(* IEC 61131-3 sources: nautilus/examples/it-rack, 2 files *)

(* ---- hw_types.st ---- *)
(*
  Generated by `naut prometheus import`: the IT-hardware UDT set from
  docs/design/it-drivers.md §2. Do not edit — every importer (snmp, redfish,
  prometheus) writes this same file, so re-running any of them restores it.
  Member order is the wire order the drivers deliver; the compiled TYPE
  must match it slot for slot, which is why it is generated and not typed.
*)

TYPE
  CPU : STRUCT
    Model : STRING;
    Cores : DINT;
    Health : DINT;
    Fault : BOOL;
    TempC : REAL;
    Pct : REAL;
  END_STRUCT;
  DIMM : STRUCT
    Locator : STRING;
    CapacityGB : REAL;
    Manufacturer : STRING;
    PartNumber : STRING;
    Health : DINT;
    Fault : BOOL;
    TempC : REAL;
  END_STRUCT;
  Drive : STRUCT
    Bay : DINT;
    Name : STRING;
    Model : STRING;
    Serial : STRING;
    CapacityGB : REAL;
    Protocol : STRING;
    MediaType : STRING;
    Health : DINT;
    Fault : BOOL;
    PredictedFailure : BOOL;
    TempC : REAL;
    Present : BOOL;
  END_STRUCT;
  Fan : STRUCT
    Name : STRING;
    Present : BOOL;
    RPM : REAL;
    Pct : REAL;
    Fault : BOOL;
  END_STRUCT;
  NetPort : STRUCT
    Name : STRING;
    LinkUp : BOOL;
    SpeedGbps : REAL;
    MAC : STRING;
  END_STRUCT;
  PCIeDevice : STRUCT
    Slot : DINT;
    Name : STRING;
    Model : STRING;
    Manufacturer : STRING;
    Firmware : STRING;
    Health : DINT;
    Fault : BOOL;
    Ports : DINT;
    TempC : REAL;
  END_STRUCT;
  PDU : STRUCT
    Online : BOOL;
    Name : STRING;
    Model : STRING;
    Serial : STRING;
    Amps : REAL;
    Watts : REAL;
    Overload : BOOL;
    OutletCount : DINT;
  END_STRUCT;
  PDUOutlet : STRUCT
    Index : DINT;
    Name : STRING;
    On : BOOL;
    Amps : REAL;
    Watts : REAL;
  END_STRUCT;
  PSU : STRUCT
    Name : STRING;
    Present : BOOL;
    Fault : BOOL;
    InputOk : BOOL;
    InputV : REAL;
    OutputW : REAL;
    CapacityW : REAL;
  END_STRUCT;
  Server : STRUCT
    Online : BOOL;
    PowerOn : BOOL;
    Health : DINT;
    Fault : BOOL;
    Warning : BOOL;
    Model : STRING;
    Serial : STRING;
    UptimeS : DINT;
    CpuPct : REAL;
    MemPct : REAL;
    Load1 : REAL;
    RootDiskPct : REAL;
    InletTempC : REAL;
    MaxTempC : REAL;
    PowerW : REAL;
    FanCount : DINT;
    PsuCount : DINT;
    TempCount : DINT;
  END_STRUCT;
  Switch : STRUCT
    Online : BOOL;
    Name : STRING;
    Model : STRING;
    Serial : STRING;
    UptimeS : DINT;
    CpuPct : REAL;
    MemPct : REAL;
    TempC : REAL;
    Fault : BOOL;
    PortsTotal : DINT;
    PortsUp : DINT;
  END_STRUCT;
  SwitchPort : STRUCT
    Index : DINT;
    Name : STRING;
    Alias : STRING;
    AdminUp : BOOL;
    OperUp : BOOL;
    Down : BOOL;
    SpeedMbps : REAL;
    InBps : REAL;
    OutBps : REAL;
    InPct : REAL;
    OutPct : REAL;
    InErrors : DINT;
    OutErrors : DINT;
    InDiscards : DINT;
    OutDiscards : DINT;
    ErrorRate : REAL;
    PoeOn : BOOL;
    PoeW : REAL;
    InBroadcastPps : REAL;
    InMulticastPps : REAL;
  END_STRUCT;
  TempSensor : STRUCT
    Name : STRING;
    Value : REAL;
    Fault : BOOL;
    High : BOOL;
    HighHigh : BOOL;
    HighSP : REAL;
    HighHighSP : REAL;
  END_STRUCT;
  UPS : STRUCT
    Online : BOOL;
    Name : STRING;
    Model : STRING;
    Serial : STRING;
    OnBattery : BOOL;
    LowBattery : BOOL;
    BatteryFault : BOOL;
    Fault : BOOL;
    ChargePct : REAL;
    RuntimeMin : REAL;
    LoadPct : REAL;
    InputV : REAL;
    OutputV : REAL;
    BatteryTempC : REAL;
  END_STRUCT;
END_TYPE

(* ---- rack.st ---- *)
(* rack.st — the rollups a rack needs that no single device carries: how
   many switch ports are up, whether anything in the rack is faulted, and
   the hottest thing in it. Everything else — every port's status, every
   fan's RPM, every sensor's thresholds — is already a UDT tag the drivers
   deliver, alarmed by the rules in nautilus.yaml, so this program stays
   small on purpose.

   Every driver-fed tag is read under its source's __Online companion: a
   device that stops answering keeps its last values (Stale) rather than
   dropping to zero, so the guard is what keeps a dark switch from being
   counted as 24 healthy ports. *)
PROGRAM Rack
VAR_EXTERNAL
  SW1 : Switch;
  SW1_Port01 : SwitchPort; SW1_Port02 : SwitchPort; SW1_Port03 : SwitchPort; SW1_Port04 : SwitchPort;
  SW1_Port05 : SwitchPort; SW1_Port06 : SwitchPort; SW1_Port07 : SwitchPort; SW1_Port08 : SwitchPort;
  SW1_Port09 : SwitchPort; SW1_Port10 : SwitchPort; SW1_Port11 : SwitchPort; SW1_Port12 : SwitchPort;
  SW1_Port13 : SwitchPort; SW1_Port14 : SwitchPort; SW1_Port15 : SwitchPort; SW1_Port16 : SwitchPort;
  SW1_Port17 : SwitchPort; SW1_Port18 : SwitchPort; SW1_Port19 : SwitchPort; SW1_Port20 : SwitchPort;
  SW1_Port21 : SwitchPort; SW1_Port22 : SwitchPort; SW1_Port23 : SwitchPort; SW1_Port24 : SwitchPort;
  SW1_Port25 : SwitchPort; SW1_Port26 : SwitchPort; SW1_Port27 : SwitchPort; SW1_Port28 : SwitchPort;
  SW1__Online : BOOL;
  MIRA1 : Server;
  MIRA1__Online : BOOL;

  PortsUp : INT;
  PortsDown : INT;
  DevicesOnline : INT;
  RackFault : BOOL;
  RackMaxTempC : REAL;
END_VAR
VAR
  up : INT;
  down : INT;
END_VAR

DevicesOnline := 0;
IF SW1__Online THEN DevicesOnline := DevicesOnline + 1; END_IF;
IF MIRA1__Online THEN DevicesOnline := DevicesOnline + 1; END_IF;

(* Ports: up = link; down = enabled but no link (Down is the driver's own
   derived member, AdminUp AND NOT OperUp — a port nobody enabled is
   neither). *)
up := 0; down := 0;
IF SW1__Online THEN
  IF SW1_Port01.OperUp THEN up := up + 1; END_IF; IF SW1_Port01.Down THEN down := down + 1; END_IF;
  IF SW1_Port02.OperUp THEN up := up + 1; END_IF; IF SW1_Port02.Down THEN down := down + 1; END_IF;
  IF SW1_Port03.OperUp THEN up := up + 1; END_IF; IF SW1_Port03.Down THEN down := down + 1; END_IF;
  IF SW1_Port04.OperUp THEN up := up + 1; END_IF; IF SW1_Port04.Down THEN down := down + 1; END_IF;
  IF SW1_Port05.OperUp THEN up := up + 1; END_IF; IF SW1_Port05.Down THEN down := down + 1; END_IF;
  IF SW1_Port06.OperUp THEN up := up + 1; END_IF; IF SW1_Port06.Down THEN down := down + 1; END_IF;
  IF SW1_Port07.OperUp THEN up := up + 1; END_IF; IF SW1_Port07.Down THEN down := down + 1; END_IF;
  IF SW1_Port08.OperUp THEN up := up + 1; END_IF; IF SW1_Port08.Down THEN down := down + 1; END_IF;
  IF SW1_Port09.OperUp THEN up := up + 1; END_IF; IF SW1_Port09.Down THEN down := down + 1; END_IF;
  IF SW1_Port10.OperUp THEN up := up + 1; END_IF; IF SW1_Port10.Down THEN down := down + 1; END_IF;
  IF SW1_Port11.OperUp THEN up := up + 1; END_IF; IF SW1_Port11.Down THEN down := down + 1; END_IF;
  IF SW1_Port12.OperUp THEN up := up + 1; END_IF; IF SW1_Port12.Down THEN down := down + 1; END_IF;
  IF SW1_Port13.OperUp THEN up := up + 1; END_IF; IF SW1_Port13.Down THEN down := down + 1; END_IF;
  IF SW1_Port14.OperUp THEN up := up + 1; END_IF; IF SW1_Port14.Down THEN down := down + 1; END_IF;
  IF SW1_Port15.OperUp THEN up := up + 1; END_IF; IF SW1_Port15.Down THEN down := down + 1; END_IF;
  IF SW1_Port16.OperUp THEN up := up + 1; END_IF; IF SW1_Port16.Down THEN down := down + 1; END_IF;
  IF SW1_Port17.OperUp THEN up := up + 1; END_IF; IF SW1_Port17.Down THEN down := down + 1; END_IF;
  IF SW1_Port18.OperUp THEN up := up + 1; END_IF; IF SW1_Port18.Down THEN down := down + 1; END_IF;
  IF SW1_Port19.OperUp THEN up := up + 1; END_IF; IF SW1_Port19.Down THEN down := down + 1; END_IF;
  IF SW1_Port20.OperUp THEN up := up + 1; END_IF; IF SW1_Port20.Down THEN down := down + 1; END_IF;
  IF SW1_Port21.OperUp THEN up := up + 1; END_IF; IF SW1_Port21.Down THEN down := down + 1; END_IF;
  IF SW1_Port22.OperUp THEN up := up + 1; END_IF; IF SW1_Port22.Down THEN down := down + 1; END_IF;
  IF SW1_Port23.OperUp THEN up := up + 1; END_IF; IF SW1_Port23.Down THEN down := down + 1; END_IF;
  IF SW1_Port24.OperUp THEN up := up + 1; END_IF; IF SW1_Port24.Down THEN down := down + 1; END_IF;
  IF SW1_Port25.OperUp THEN up := up + 1; END_IF; IF SW1_Port25.Down THEN down := down + 1; END_IF;
  IF SW1_Port26.OperUp THEN up := up + 1; END_IF; IF SW1_Port26.Down THEN down := down + 1; END_IF;
  IF SW1_Port27.OperUp THEN up := up + 1; END_IF; IF SW1_Port27.Down THEN down := down + 1; END_IF;
  IF SW1_Port28.OperUp THEN up := up + 1; END_IF; IF SW1_Port28.Down THEN down := down + 1; END_IF;
END_IF;
PortsUp := up;
PortsDown := down;

(* Rack health: any device faulted, or any device dark. *)
RackFault := (SW1__Online AND SW1.Fault) OR (MIRA1__Online AND MIRA1.Fault)
             OR NOT SW1__Online OR NOT MIRA1__Online;

(* The hottest reading in the rack, over the devices that report one. *)
RackMaxTempC := 0.0;
IF SW1__Online AND SW1.TempC > RackMaxTempC THEN RackMaxTempC := SW1.TempC; END_IF;
IF MIRA1__Online AND MIRA1.MaxTempC > RackMaxTempC THEN RackMaxTempC := MIRA1.MaxTempC; END_IF;
END_PROGRAM
